FUNCTION_BLOCK BasicHashTest (* Basic FB with an ECC *)
  (* Standard: 61499-1; Description: Copyright (c) 2026 Martin Erich Jobst This program and the accompanying materials are made available under the terms of the Eclipse Public License 2.0 which is available at https://www.eclipse.org/legal/epl-2.0/ SPDX-License-Identifier: EPL-2.0 *)
  (* Version 1.0, 2026-10-28, Martin Jobst *)
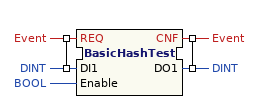
  EVENT_INPUT
    REQ WITH DI1; (* Request *)
  END_EVENT
  EVENT_OUTPUT
    CNF WITH DO1; (* Confirmation *)
  END_EVENT
  VAR_INPUT
    DI1 : DINT := DINT#1;
    Enable : BOOL := TRUE;
  END_VAR
  VAR_OUTPUT
    DO1 : DINT := DINT#0;
  END_VAR
  VAR CONSTANT
    limit : DINT := DINT#10;
  END_VAR
  VAR
    counter : DINT := DINT#0;
  END_VAR
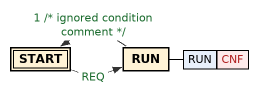
  EC_STATES
    START; (* Initial State *)
    RUN : RUN -> CNF;
  END_STATES
  EC_TRANSITIONS
    START TO RUN := REQ;
    RUN TO START := 1 /* ignored condition comment */;
  END_TRANSITIONS
  ALGORITHM RUN IN ST:
	IF Enable THEN
		counter := counter + DI1;
	END_IF;
	DO1 := MIN(counter, limit);
  END_ALGORITHM
END_FUNCTION_BLOCK
